// TIA Portal V14 SP1 export
// export: Created 2000-01-01T00:00:00.0000000Z, ExportSetting None
FUNCTION "MCP_RC_FCmin" : Void   // FC9810, LAD
{ S7_Optimized_Access := 'TRUE' }
   VAR_INPUT
      "A" : Bool;
   END_VAR
BEGIN
END_FUNCTION
